(* IEC 61131-3 sources: repolevel_ST_code_completion/ground_truth/repoeval_four-level_elevator_control/readful_result, 2 files *)

(* ---- F_CheckJobInDirection.st ---- *)
It seems like you've provided a code fragment for a function named `F_CheckJobInDirection` written in Structured Text (ST), which is commonly used in PLC programming. The function checks whether there are any elevator stop requests between two floors (`nStartFloor` and `nEndFloor`) in a specified direction (`bIncreasing`).

However, the code fragment appears to be incomplete or repeated multiple times. Below is a cleaned-up and complete version of the function based on the provided snippets:

```pascal
FUNCTION F_CheckJobInDirection : BOOL
VAR_INPUT
	nStartFloor		:	USINT;		// 起始楼层
	nEndFloor		:	USINT;		// 结束楼层
	bIncreasing		:	BOOL;		// TRUE=向上检查（递增），FALSE=向下检查（递减）
END_VAR
VAR
	i	:	USINT;	// 循环变量
END_VAR

// 初始化返回值为 FALSE
F_CheckJobInDirection := FALSE;

IF bIncreasing THEN
	// 向上检查（从低楼层到高楼层）
	FOR i := nStartFloor TO nEndFloor DO
		IF Tar_Dir.IsStopFloor[i] THEN
			F_CheckJobInDirection := TRUE;
			RETURN; // 如果找到需要停靠的楼层，立即返回 TRUE
		END_IF
	END_FOR
ELSE
	// 向下检查（从高楼层到低楼层）
	FOR i := nEndFloor TO nStartFloor BY -1 DO
		IF Tar_Dir.IsStopFloor[i] THEN
			F_CheckJobInDirection := TRUE;
			RETURN; // 如果找到需要停靠的楼层，立即返回 TRUE
		END_IF
	END_FOR
END_IF
```

### Explanation of the Code:
1. **Inputs**:
   - `nStartFloor`: The starting floor for the check.
   - `nEndFloor`: The ending floor for the check.
   - `bIncreasing`: A boolean indicating the direction of the check (`TRUE` for upward, `FALSE` for downward).

2. **Logic**:
   - If `bIncreasing` is `TRUE`, the function iterates from `nStartFloor` to `nEndFloor` (low to high).
   - If `bIncreasing` is `FALSE`, the function iterates from `nEndFloor` to `nStartFloor` (high to low).
   - During each iteration, it checks if the current floor (`i`) is marked as a stop floor (`Tar_Dir.IsStopFloor[i]`).
   - If a stop floor is found, the function sets the return value to `TRUE` and exits immediately using `RETURN`.

3. **Return Value**:
   - The function returns `TRUE` if there is at least one stop floor in the specified range and direction.
   - Otherwise, it returns `FALSE`.

### Notes:
- The variable `Tar_Dir.IsStopFloor` is assumed to be an array or similar data structure that indicates whether a specific floor is a stop floor.
- Ensure that the indices for `Tar_Dir.IsStopFloor` are valid and within bounds to avoid runtime errors.
- The function is designed to be efficient by exiting as soon as a stop floor is found.

If you have additional questions or need further clarification, feel free to ask!

(* ---- F_CheckJobInDirection_1.st ---- *)
It seems like you've provided a code fragment for a function named `F_CheckJobInDirection` written in Structured Text (ST), which is commonly used in PLC programming. The function checks whether there are any elevator stop requests between two floors (`nStartFloor` and `nEndFloor`) in a specified direction (`bIncreasing`).

However, the code fragment appears to be incomplete or repeated multiple times. Below is a cleaned-up and complete version of the function based on the provided snippets:

```pascal
FUNCTION F_CheckJobInDirection : BOOL
VAR_INPUT
	nStartFloor		:	USINT;		// 起始楼层
	nEndFloor		:	USINT;		// 结束楼层
	bIncreasing		:	BOOL;		// TRUE=向上检查（递增），FALSE=向下检查（递减）
END_VAR
VAR
	i	:	USINT;	// 循环变量
END_VAR

// 初始化返回值为 FALSE
F_CheckJobInDirection := FALSE;

IF bIncreasing THEN
	// 向上检查（从低楼层到高楼层）
	FOR i := nStartFloor TO nEndFloor DO
		IF Tar_Dir.IsStopFloor[i] THEN
			F_CheckJobInDirection := TRUE;
			RETURN; // 如果找到需要停靠的楼层，立即返回 TRUE
		END_IF
	END_FOR
ELSE
	// 向下检查（从高楼层到低楼层）
	FOR i := nEndFloor TO nStartFloor BY -1 DO
		IF Tar_Dir.IsStopFloor[i] THEN
			F_CheckJobInDirection := TRUE;
			RETURN; // 如果找到需要停靠的楼层，立即返回 TRUE
		END_IF
	END_FOR
END_IF
```

### Explanation of the Code:
1. **Inputs**:
   - `nStartFloor`: The starting floor for the check.
   - `nEndFloor`: The ending floor for the check.
   - `bIncreasing`: A boolean indicating the direction of the check (`TRUE` for upward, `FALSE` for downward).

2. **Logic**:
   - If `bIncreasing` is `TRUE`, the function iterates from `nStartFloor` to `nEndFloor` (low to high).
   - If `bIncreasing` is `FALSE`, the function iterates from `nEndFloor` to `nStartFloor` (high to low).
   - During each iteration, it checks if the current floor (`i`) is marked as a stop floor (`Tar_Dir.IsStopFloor[i]`).
   - If a stop floor is found, the function sets the return value to `TRUE` and exits immediately using `RETURN`.

3. **Return Value**:
   - The function returns `TRUE` if there is at least one stop floor in the specified range and direction.
   - Otherwise, it returns `FALSE`.

### Notes:
- The variable `Tar_Dir.IsStopFloor` is assumed to be an array or similar data structure that indicates whether a specific floor is a stop floor.
- Ensure that the indices for `Tar_Dir.IsStopFloor` are valid and within bounds to avoid runtime errors.
- The function is designed to be efficient by exiting as soon as a stop floor is found.

If you have additional questions or need further clarification, feel free to ask!
